(*
SPDX-FileCopyrightText: © 2026 Oleksandr Tiutyk <trofimich@gmail.com>
SPDX-License-Identifier: MIT
License: https://opensource.org/license/mit
*)

(*!
<summary>Reports a field or property whose TwinCAT type class is unsupported.</summary>
<description>
The caller detects the member error; Throw records diagnostics rather than inspecting the object. Dynamic
instances and clones belong to the current task memory manager until cleanup. Dynamic copies are explicitly
registered by Clone after construction; plain __NEW does not transfer ownership to the task manager.
Runtime type diagnostics use TYPE_ names for known classes and decimal codes for unknown values.
</description>
*)

{attribute 'enable_dynamic_creation'}
{attribute 'no_explicit_call' := 'do not call this function block directly'}
FUNCTION_BLOCK DataMemberTypeClassNotSupportedException EXTENDS GeneralException IMPLEMENTS IDataMemberTypeClassNotSupportedException
VAR_STAT
	//! <summary>Class name shared by all instances of this function block.</summary>
	{attribute 'hide'} 
	_ClassName : STRING := __POUNAME();
END_VAR

{attribute 'monitoring' := 'call'}
PROPERTY ClassName : REFERENCE TO STRING
GET
ClassName REF= _ClassName;
END_GET
END_PROPERTY

(*!
<summary>Creates a distinct auto-disposed copy of this concrete exception type.</summary>
<description>
Copies message, code, source and timestamps through CopyGeneralFields; any prepared inner cause remains
borrowed. The current task memory manager owns the clone until cleanup. Allocation failure is terminal.
Descendants with additional payload must override Clone to preserve their type and fields. Registers the newly
constructed instance before copying payload, outside FB_init. Registration failure releases the unregistered
instance and raises a terminal error; copy failure leaves the registered instance owned by the task manager
for cleanup. Custom overrides must follow the same ownership sequence.
</description>
*)
METHOD Clone : IObject
VAR
	exceptionClone : POINTER TO DataMemberTypeClassNotSupportedException;
END_VAR
exceptionClone := __NEW(DataMemberTypeClassNotSupportedException);

IF exceptionClone = 0 THEN
	DynamicMemoryManager.RaiseAllocationFailure();
END_IF

DynamicMemoryManager.RegisterAutoDisposedObject(autoDisposedObject := exceptionClone^);

exceptionClone^.CopyGeneralFields(sourceException := THIS^);

Clone := exceptionClone^;
END_METHOD

(*!
<summary>Provides the library namespace used in diagnostics.</summary>
<description>
Borrowed read-only reference to the compiler-initialized library namespace; no ownership transfer.
</description>
*)
{attribute 'monitoring' := 'call'}
PROPERTY NamespaceName : REFERENCE TO STRING
GET
NamespaceName REF= CurrentNamespace.Name;
END_GET
END_PROPERTY

(*!
<summary>Reports the byte size of this concrete instance.</summary>
<description>
Uses XSIZEOF on the instance. Does not include separately allocated payloads or prove that an arbitrary
address is valid.
</description>
*)
{attribute 'monitoring' := 'call'}
PROPERTY SelfSize : ULINT
GET
SelfSize := XSIZEOF(THIS^);
END_GET
END_PROPERTY

(*!
<summary>Formats the rejected member and propagates the exception.</summary>
<description>
Call in the owning cyclic task, not during FB_init. Builds a member diagnostic without heap allocation during
message preparation and captures source and timestamps with zero error code and no inner cause. Input storage
is not retained. Exception clone allocation failure uses the shared terminal memory mechanism.
Known runtime type classes appear by their TYPE_ names; unknown values retain their decimal codes.
</description>
<param name="dataMemberName">Name of the field or property rejected by the caller.</param>
<param name="dataMemberType">Unsupported TwinCAT type class.</param>
*)
METHOD Throw
VAR_INPUT
	sourceNamespaceName : STRING;
	sourceClassName : STRING;
	sourcePOUName : STRING;
	sourcePosition : STRING;
	dataMemberName : STRING;
	dataMemberType : __SYSTEM.TYPE_CLASS;
END_VAR
VAR
	message : ERROR_MESSAGE;
END_VAR
WideStrings.Append255(
	message,
	"Field or property '",
	TO_WSTRING(dataMemberName),
	"' has not supported type class '",
	SystemTypeClassConvertor.ToWideString(typeClass := dataMemberType),
	"' in the instance of '",
	TO_WSTRING(sourceNamespaceName),
	".",
	TO_WSTRING(sourceClassName),
	"'");

InternalThrow(
	sourceNamespaceName := sourceNamespaceName,
	sourceClassName := sourceClassName,
	sourcePOUName := sourcePOUName,
	sourcePosition := sourcePosition,
	message := message,
	errorCode := 0,
	innerException := 0
);
END_METHOD

END_FUNCTION_BLOCK

(* stored: Version 1.1.0.1
   POU DataMemberTypeClassNotSupportedException: Id {61dbf5b4-4beb-4336-96b1-4503e29de50d}, SpecialFunc None
   Property ClassName: Id {a3aa58b0-7b00-447c-9463-7b40f3db7b6d}
   Get Get: Id {225dea7c-7ed1-4b1b-9aa9-e37bc958cb35}
   Method Clone: Id {5fce08bb-c660-4608-89d3-b9d6be39bbc0}
   Property NamespaceName: Id {5eb62e43-021c-4874-a255-47e07f04825b}
   Get Get: Id {af49da20-ade9-4011-9b13-bad8b4fbc737}
   Property SelfSize: Id {c7958ef8-cf29-412d-b3ad-0101df0c5c1a}
   Get Get: Id {7b643129-d919-4326-bde2-8d1483b19251}
   Method Throw: Id {f1d83160-3a5d-4dd9-a889-f5f3673452d9} *)
